Fanuc TP program (LS listing): EdgePr.LS

/PROG  EdgePr
/ATTR
OWNER		= MNEDITOR;
COMMENT		= "RoboDK sequence";
PROG_SIZE	= 0;
CREATE		= DATE 31-12-14  TIME 12:00:00;
MODIFIED	= DATE 31-12-14  TIME 12:00:00;
FILE_NAME	= EdgePr;
VERSION		= 0;
LINE_COUNT	= 39;
MEMORY_SIZE	= 0;
PROTECT		= READ_WRITE;
TCD:  STACK_SIZE	= 0,
      TASK_PRIORITY	= 50,
      TIME_SLICE	= 0,
      BUSY_LAMP_OFF	= 0,
      ABORT_REQUEST	= 0,
      PAUSE_REQUEST	= 0;
DEFAULT_GROUP	= 1,*,*,*,*;
CONTROL_CODE	= 00000000 00000000;
/MN
   1:  ! Program generated by RoboDK v6.0.7 for Fanuc ARC Mate 100iD/8 ;
   2:  ! L on XX/XX/XXXX 18:00:00 ;
   3:  ! Using nominal kinematics. ;
   4:  PR[9,1]=100.500 ;
   5:  PR[9,2]=-200.250 ;
   6:  PR[9,3]=300.125 ;
   7:  PR[9,4]=30.000 ;
   8:  PR[9,5]=-20.000 ;
   9:  PR[9,6]=10.000 ;
  10:  UFRAME[9]=PR[9] ;
  11:  UFRAME_NUM=9 ;
  12:  PR[9,1]=-1.500 ;
  13:  PR[9,2]=2.250 ;
  14:  PR[9,3]=99.875 ;
  15:  PR[9,4]=180.000 ;
  16:  PR[9,5]=45.000 ;
  17:  PR[9,6]=-90.000 ;
  18:  UTOOL[9]=PR[9] ;
  19:  UTOOL_NUM=9 ;
  20:J P[1] 17% FINE ;
  21:L P[2] 123mm/sec CNT12 ;
  22:  PAUSE ;
  23:  WAIT  1.23(sec) ;
  24:  MESSAGE[A long message with "quotes", 'apostrophes' & symbols:] ;
  25:  MESSAGE[<>[]{}()=+-*/%;#@! and more text to make it longer th] ;
  26:  MESSAGE[an eighty characters] ;
  27:  ! Comment with ; semicolon ;
  28:  Gripper=(ON) ;
  29:  DO[12]=OFF ;
  30:  Pressure=(0.75) ;
  31:  $WAITTMOUT=250 ;
  32:  WAIT PartPresent=ON TIMEOUT, LBL[1] ;
  33:  MESSAGE[Timed out for LBL 1] ;
  34:  PAUSE ;
  35:  LBL[1] ;
  36:  WAIT DI[7]=(1) ;
  37:  CALL DoSometh(1, 2) ;
  38:  x = 1;
  39:J P[3] 17% CNT12 ;
/POS
P[1]{
   GP1:
    UF : 9, UT : 9,
	J1=    -5.000 deg,	J2=    -5.000 deg,	J3=    15.000 deg,
	J4=    10.000 deg,	J5=    40.000 deg,	J6=    -10.000 deg
};
P[2]{
   GP1:
    UF : 9, UT : 9,        CONFIG : 'F U T, 0, 0, 0',
	X =  -624.230  mm,	Y =   571.208  mm,	Z =   454.620  mm,
	W =   -82.711 deg,	P =    44.567 deg,	R =  -122.815 deg
};
P[3]{
   GP1:
    UF : 9, UT : 9,
	J1=    20.000 deg,	J2=    -10.000 deg,	J3=    20.000 deg,
	J4=    0.000 deg,	J5=    30.000 deg,	J6=    0.000 deg
};
/END
